Universal Robots URScript: letra_J.script

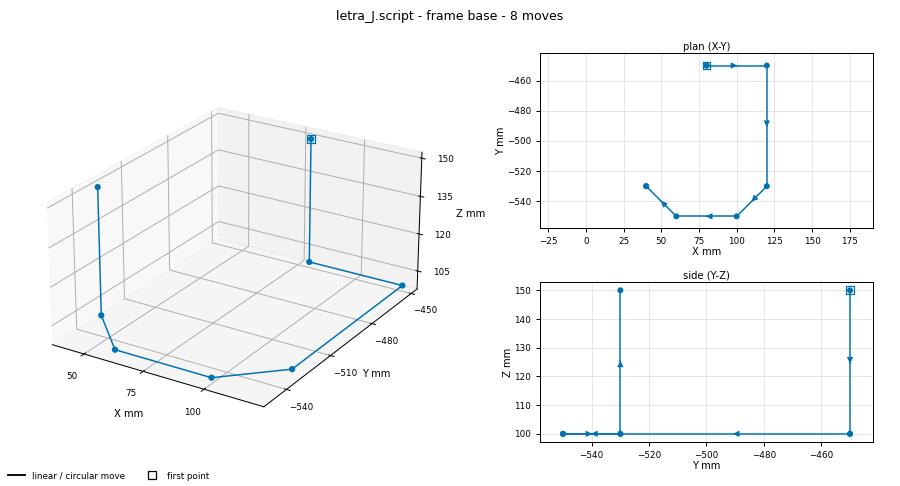
[picture p0: tool path of letra_J.script in frame base, 8 of 8 moves have a stored position in this frame; points joined in program order, loops and branches not executed]
# Letra J - Juan
movel(p[0.080, -0.450, 0.150, 3.1416, 0, 0], a=0.5, v=0.1)
movel(p[0.080, -0.450, 0.100, 3.1416, 0, 0], a=0.5, v=0.1)
movel(p[0.120, -0.450, 0.100, 3.1416, 0, 0], a=0.5, v=0.1)
movel(p[0.120, -0.530, 0.100, 3.1416, 0, 0], a=0.5, v=0.1)
movel(p[0.100, -0.550, 0.100, 3.1416, 0, 0], a=0.5, v=0.1)
movel(p[0.060, -0.550, 0.100, 3.1416, 0, 0], a=0.5, v=0.1)
movel(p[0.040, -0.530, 0.100, 3.1416, 0, 0], a=0.5, v=0.1)
movel(p[0.040, -0.530, 0.150, 3.1416, 0, 0], a=0.5, v=0.1)
